FUNCTION_BLOCK GATE_CYCLE
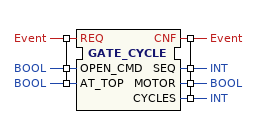
  EVENT_INPUT
    REQ WITH OPEN_CMD, AT_TOP;
  END_EVENT
  EVENT_OUTPUT
    CNF WITH SEQ, MOTOR, CYCLES;
  END_EVENT
  VAR_INPUT
    OPEN_CMD : BOOL;
    AT_TOP : BOOL;
  END_VAR
  VAR_OUTPUT
    SEQ : INT;
    MOTOR : BOOL;
    CYCLES : INT;
  END_VAR
  VAR
    K : INT;
  END_VAR
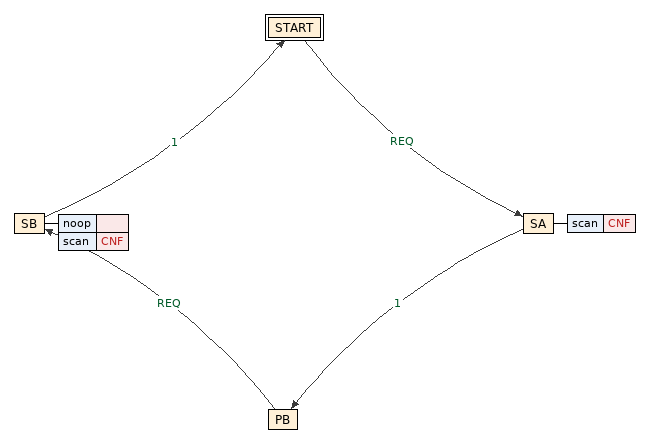
  EC_STATES
    START;
    SA : scan -> CNF;
    PB;
    SB : noop, scan -> CNF;
  END_STATES
  EC_TRANSITIONS
    START TO SA := REQ;
    SA TO PB := 1;
    PB TO SB := REQ;
    SB TO START := 1;
  END_TRANSITIONS
  ALGORITHM scan IN ST:
K := SEQ;
MOTOR := FALSE;
CASE K OF
 0: IF OPEN_CMD THEN SEQ := 1; END_IF;
 1: MOTOR := TRUE; IF AT_TOP THEN SEQ := 2; END_IF;
 2: CYCLES := CYCLES + 1; SEQ := 0;
END_CASE;
  END_ALGORITHM
  ALGORITHM noop IN ST:
K := 0;
  END_ALGORITHM
END_FUNCTION_BLOCK
